Fanuc KAREL source: KO00004.KL

PROGRAM KO00004
%NOLOCKGROUP
VAR
  P1: POSITION
  P2: POSITION
  P3: POSITION
  OUT: JOINTPOS
BEGIN
  OUT = FRAME(P1, P2, P3)
END KO00004
